Staubli VAL3: refreshlist.pgx

public program refreshlist()
  local string l_skey
  local num l_i
  local num l_nSize
begin
  call program:getProgList(sProgLsit)
  l_nSize=size(sProgLsit)

  if l_nSize<=49
    nPageNum=1
  else
    nPageNum=roundUp(l_nSize/49)
  endIf

  if nPageNum==1
    for l_i = 0 to size(sList)-1
      sList[l_i]=""
    endFor
    for l_i = 0 to l_nSize-1
      sList[l_i]=sProgLsit[l_i]
    endFor
  else
    if nPageIndex<nPageNum-1
      for l_i = 0 to 48
        sList[l_i]=sProgLsit[49*nPageIndex+l_i]
      endFor
    else
      for l_i = 0 to size(sList)-1
        sList[l_i]=""
      endFor
      for l_i = 0 to(l_nSize%49)-1
        sList[l_i]=sProgLsit[49*nPageIndex+l_i]
      endFor
    endIf
  endIf
  userPageBind("prog","lst1","options",sList,size(sList),"r")
  sPageIndex=toString("",nPageIndex+1)
  sPageNum=toString("",nPageNum)
end
